Universal Robots URScript: T006_mistralai_Devstral-Small-2-24B-Instruct-2512_baseline_rep1_retry2.urscript

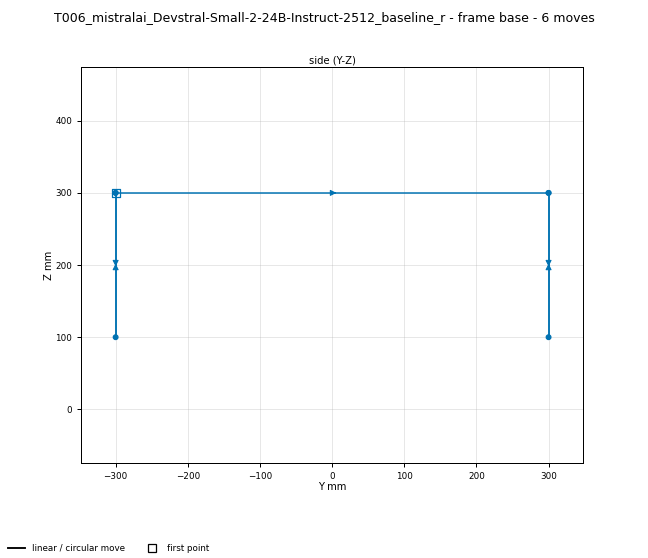
[picture p0: tool path of T006_mistralai_Devstral-Small-2-24B-Instruct-2512_baseline_rep1_retry2.urscript in frame base, 6 of 8 moves have a stored position in this frame; points joined in program order, loops and branches not executed]
def bin_picking_suction():
    # Home position
    movej([0, -1.5708, 0, -1.5708, -1.5708, 0], a=350.0, v=350.0)

    # Above bin
    tool_on()
    movel(p[0.5, -0.3, 0.3, 0, 3.1416, 0], a=350.0, v=350.0)

    # Descend into bin
    movel(p[0.5, -0.3, 0.1, 0, 3.1416, 0], a=150.0, v=150.0)

    # Lift from bin
    movel(p[0.5, -0.3, 0.3, 0, 3.1416, 0], a=300.0, v=300.0)

    # Transit to conveyor
    movel(p[0.5, 0.3, 0.3, 0, 3.1416, 0], a=380.0, v=380.0)

    # Descend to conveyor
    movel(p[0.5, 0.3, 0.1, 0, 3.1416, 0], a=300.0, v=300.0)

    # Release part
    tool_off()
    sleep(1.0)

    # Lift from conveyor
    movel(p[0.5, 0.3, 0.3, 0, 3.1416, 0], a=300.0, v=300.0)

    # Return to home
    movej([0, -1.5708, 0, -1.5708, -1.5708, 0], a=350.0, v=350.0)

    # End program
    end_program()
